// TIA Portal V20 export
// export: Created 2026-10-19T18:41:42.5052307Z, ExportSetting WithDefaults, DisplayName Totally Integrated Automation Portal, DisplayVersion V20 Update 6, DisplayName TIA Portal Openness, DisplayVersion V20 Update 6, DisplayName TIA Portal Version Control Interface, DisplayVersion V20 Update 6, DisplayName SINAMICS Startdrive Advanced, DisplayVersion V20 SP1, DisplayName SINAMICS Startdrive G130, G150, S120, S150, SINAMICS MV, G220, S200, S210, DisplayVersion V20 SP1, DisplayName SINAMICS Startdrive G110M, G120, G120C, G120D, G120P, G115D, DisplayVersion V20 SP1, DisplayName STEP 7 Professional, DisplayVersion V20 Update 6, DisplayName STEP 7 Safety, DisplayVersion V20 Update 2, DisplayName WinCC Basic/Comfort/Advanced, DisplayVersion V20 Update 6, DisplayName WinCC Unified, DisplayVersion V20 Update 6
DATA_BLOCK "FB_HeartBeat_DB"   // DB136
VERSION : 0.1
// stored: AutoNumber true, DBAccessibleFromOPCUA true, InstanceOfName FB_HeartBeat, InstanceOfType FB
"FB_HeartBeat"
   // VAR_INPUT
   //    PC_HeartBeat : Word := 16#6E87;
   // END_VAR
   // VAR_OUTPUT
   //    PLC_HeartBeat : Word := 16#B1B0;
   //    PC_Disconnected : Bool := TRUE;
   // END_VAR
   // VAR
   //    TimeOut : TON_TIME;
   //    "Timer" { S7_SetPoint := 'True'} : TON_TIME;
   //    PC_Heartbeat_old : Word := 16#6E87;
   //    StartTimerBit : Bool;
   // END_VAR
BEGIN
   TimeOut.PT := T#10S;
   TimeOut.IN := TRUE;
   "Timer".PT := T#500MS;
   "Timer".IN := TRUE;
END_DATA_BLOCK
